TYPE ST_BeadUp :
STRUCT
	lrBeadUpForce						:LREAL;											(* BeadUp force [N] *)
	unBeadUpRamp						:UINT;											(* BeadUp ramp [s] *)
	unBeadUpTime						:UINT;											(* BeadUp time [s] *)
	lrVeloForceCtrlKp						:LREAL;											(* Velocity - force controller proportional band Kp *)
	lrVeloForceCtrlTi						:LREAL;											(* Velocity - force controller integral Ti *)
	lrVeloForceCtrlLimit					:LREAL;											(* Velocity - force controller limit  *)
END_STRUCT
END_TYPE

(* stored: Version 1.1.0.1, ProductVersion 3.1.4024.15
   DUT ST_BeadUp: Id {fff0d6af-4c9c-4b1b-957c-e9aa89f6e25e} *)
